Fanuc KAREL source: kd00003.KL

PROGRAM KD00003
%STACKSIZE=65535
%PRIORITY=65535
%CMOSVARS
%NOLOCKGROUP
VAR
I : INTEGER
J : INTEGER
B : BOOLEAN
R : REAL
S : STRING[80]
BEGIN
I=1
END KD00003
